(* IEC 61131-3 sources: codesys-to-s7/tests/corpus/C2S7-SEM-CTR/pos, 1 file *)

(* ---- input.st ---- *)
FUNCTION_BLOCK FB_Case
VAR
    c : CTU;
    x : BOOL;
END_VAR
c(CU := x, PV := 10);
END_FUNCTION_BLOCK
